(* IEC 61131-3 sources: volt/packages/volt-lsp-iec/test-corpus/CodesysTestProject/Device/Plc Logic/Application, 3 files *)

(* ---- VltFixtureCfc.pou ---- *)
FUNCTION_BLOCK VltFixtureCfc
VAR_INPUT
END_VAR
VAR_OUTPUT
END_VAR
VAR
END_VAR

%LANGUAGE CFC UNSUPPORTED

END_FUNCTION_BLOCK

(* ---- VltFixtureSfc.pou ---- *)
FUNCTION_BLOCK VltFixtureSfc
VAR_INPUT
END_VAR
VAR_OUTPUT
END_VAR
VAR
END_VAR

%LANGUAGE SFC UNSUPPORTED

END_FUNCTION_BLOCK

(* ---- PLC_PRG.pou ---- *)
PROGRAM PLC_PRG
VAR
END_VAR
%LANGUAGE ST

END_PROGRAM
